Fanuc KAREL source: KT00950.KL

PROGRAM KT00950
%NOLOCKGROUP
VAR
  ENTRY: INTEGER
  PNAME: STRING[80]
  VNAME: STRING[80]
  STATUS: INTEGER
  VALUE: ARRAY[4] OF SHORT
BEGIN
  ENTRY = 0
  PNAME = ''
  VNAME = 'VALUE'
  GET_VAR(ENTRY, PNAME, VNAME, VALUE, STATUS)
END KT00950
